Universal Robots URScript: T001_qwen2.5-coder_32b-instruct-q4_0_safety_rep1.urscript

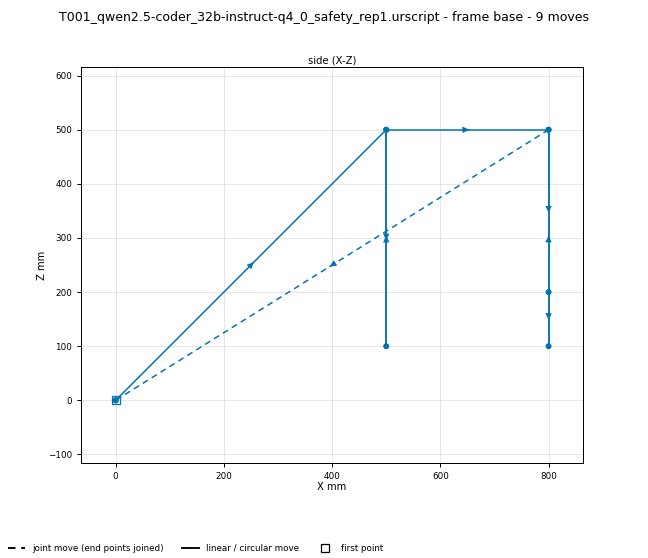
[picture p0: tool path of T001_qwen2.5-coder_32b-instruct-q4_0_safety_rep1.urscript in frame base, 9 of 9 moves have a stored position in this frame; points joined in program order, loops and branches not executed]
def safety_check():
    if not is_within_safety_zone(get_tcp_pose()):
        popup("Safety violation detected! Halting operation.")
        halt()

def is_within_safety_zone(tcp_pose):
    # Define safety zone boundaries (example values, adjust as necessary)
    x_min = -1000
    x_max = 1000
    y_min = -1000
    y_max = 1000
    z_min = 0
    z_max = 1500

    x = tcp_pose[0]
    y = tcp_pose[1]
    z = tcp_pose[2]

    return x >= x_min and x <= x_max and y >= y_min and y <= y_max and z >= z_min and z <= z_max

def main():
    set_payload(0.5, [0, 0, 0.05])

    # Home position
    safety_check()
    movej(p[0.0, -1.57, 0.0, -1.57, 0.0, 0.0], a=1.4, v=2.0)  # Adjusted to max joint acceleration

    # Approach pick point
    safety_check()
    movel(p[0.5, -1.57, 0.5, -1.57, 0.0, 0.0], a=1.4, v=2.0)  # Adjusted to max joint acceleration

    # Descend to pick
    safety_check()
    movel(p[0.5, -1.57, 0.1, -1.57, 0.0, 0.0], a=1.4, v=0.15)  # Adjusted to max joint acceleration

    # Lift from pick
    safety_check()
    movel(p[0.5, -1.57, 0.5, -1.57, 0.0, 0.0], a=1.4, v=0.1875)  # Adjusted to max joint acceleration

    # Transit to place approach
    safety_check()
    movel(p[0.8, -1.57, 0.5, -1.57, 0.0, 0.0], a=1.4, v=2.0)  # Adjusted to max joint acceleration

    # Approach place point
    safety_check()
    movel(p[0.8, -1.57, 0.2, -1.57, 0.0, 0.0], a=1.4, v=2.0)  # Adjusted to max joint acceleration

    # Descend to place
    safety_check()
    movel(p[0.8, -1.57, 0.1, -1.57, 0.0, 0.0], a=1.4, v=0.15)  # Adjusted to max joint acceleration

    # Lift from place
    safety_check()
    movel(p[0.8, -1.57, 0.5, -1.57, 0.0, 0.0], a=1.4, v=0.1875)  # Adjusted to max joint acceleration

    # Return to home
    safety_check()
    movej(p[0.0, -1.57, 0.0, -1.57, 0.0, 0.0], a=1.4, v=2.0)  # Adjusted to max joint acceleration

main()
